(* IEC 61131-3 sources: volt/packages/volt-lsp-iec/test-corpus/bakon-nano/Device/Plc Logic/Application/Library Manager/CAA Tick, 5 files *)

(* ---- PROPERTYCONSTANTS.gvl ---- *)
VAR_GLOBAL
	GC_WRESEXP : WORD := 1;
	GC_WRESNUM : WORD := 2;
	GC_WRESDENOM : WORD := 3;
	GC_WMAXINTERVAL : WORD := 10;
END_VAR

(* ---- VERSIONCONSTANTS.gvl ---- *)
VAR_GLOBAL
	GC_BYVERSION : BYTE := 1;
	GC_VERSION_1 : BYTE := 0;
END_VAR

(* ---- GETPROPERTY.pou ---- *)
FUNCTION GETPROPERTY : __XWORD
VAR_INPUT
	WPROPERTY : WORD;
END_VAR
END_FUNCTION

(* ---- GETSUPPLIERVERSION.pou ---- *)
FUNCTION GETSUPPLIERVERSION : WORD
VAR_INPUT
	XDUMMY : BOOL;
END_VAR
END_FUNCTION

(* ---- GETTICK.pou ---- *)
FUNCTION GETTICK : CAA.TICK
VAR_INPUT
	XDUMMY : BOOL;
END_VAR
END_FUNCTION
